(* IEC 61131-3 sources: ironplc/compiler/syntax/tests/fixtures/lexical, 3 files *)

(* ---- oscat_marker_in_string.st ---- *)
PROGRAM OscatMarkerInString
VAR
    text : STRING[40];
    count : INT;
END_VAR
text := '(*@KEY@:X*)';
count := count + 1;
text := '(*@KEY@:END_X*)';
END_PROGRAM

(* ---- oscat_several_pairs.st ---- *)
PROGRAM OscatSeveralPairs
(*@KEY@:DESCRIPTION*)
first documentation block, free text: it's not code ? { (*
(*@KEY@:END_DESCRIPTION*)
VAR
    count : INT;
END_VAR
(*@KEY@:NOTES*)
second documentation block, free text: it's not code ? { (*
(*@KEY@:END_NOTES*)
count := count + 1;
(*@KEY@:REVISION*)
third documentation block, `unterminated "quote
(*@KEY@:END_REVISION*)
END_PROGRAM

(* ---- unicode_comments_pragmas.st ---- *)
{attribute 'strict'}
PROGRAM Lexical	(* tab before this comment *)
VAR
	name : STRING[16]; (* café (* nested *) tab	here *)
	Größe : INT;  // line comment with ünïcode
	flag AT %IX0.0 : BOOL; /// doc comment
END_VAR
{attribute 'hide'}
name := 'Wärme $L $41';
Größe := 1;
/* block comment */ flag := TRUE;
END_PROGRAM
